FUNCTION fun_Real_SecondsToTime : TIME
VAR_INPUT
	in_Time: REAL; // Seconds

END_VAR
VAR
END_VAR

fun_Real_SecondsToTime:=DINT_TO_TIME(TRUNC(in_Time*1000));

END_FUNCTION

(* stored: Version 1.1.0.1, ProductVersion 3.1.4024.12
   POU fun_Real_SecondsToTime: Id {5e3bb995-b01d-479b-ba4a-51b69096b726}, SpecialFunc None *)
